Staubli VAL3: main.pgx

public program main(frame& x_fCellule)
  local num l_nRef0
  local num l_nResult
begin


  link(fWorld0,x_fCellule)
  l_nRef0 =0
  fWorld0.trsf = $Xposition(world,x_fCellule,l_nRef0)

  if prog:libLoad("./PROG1_withaverylongnameandspecialcharacters")!=0
    logMsg("Error Loading RoboDK library")
    popUpMsg("Error Loading RoboDK library")
  endIf
  wait(taskStatus("loading")==-1)
  prog:fPartReal.trsf=fPartCad.trsf*fCadToReal.trsf
  prog:tCad.trsf=tCad.trsf*tAdjust.trsf
  call prog:setLink(fWorld0)
  call prog:start()



end
